SUBAPPLICATION AX_TO_QXA_BG_PUBLISH (* Treibt aus einem bereits fertigen AX-Zustand (z.B. per OR mehrerer Quellen zusammengefuehrt - gestaffeltes Gruppensignal, Einzel-Toggle, IO-Diag-Testbutton) 1 physischen Ausgang + Hintergrundfarbe (SoftKey+AUX) + lokalen State-Publish (Web-Client/OPC-Dashboard). Gegenstueck zu MyLib::sys::AX_SoftkeyToggle_RS_TO_QXA_BG (das den Toggle/Reset noch selbst erzeugt) - hier liegt der AX-Zustand bereits fertig vor und muss nur noch auf Ausgang+Hintergrund+Publish verteilt werden. *)
  (* Standard: 61499-2; Description: Copyright (c) 2026 Meisterschulen am Ostbahnhof This program and the accompanying materials are made available under the terms of the Eclipse Public License 2.0 which is available at https://www.eclipse.org/legal/epl-2.0/ SPDX-License-Identifier: EPL-2.0 *)
  (* Version 1.2, 2026-10-13, Franz Höpfinger, Meisterschulen am Ostbahnhof, Neuer SubAppEventOutput INITO (Type EInit), durchgereicht von DigitalOutput.INITO - analog ILOCK_SWITCH_2_QXA_OPC v1.3, fuer die Option-Lib-Migration Igel/Elevator Klassisch (echtes INIT_CNF statt T#15s-Delay-Raten). *)
  (* Version 1.1, 2026-10-12, Franz Höpfinger, Meisterschulen am Ostbahnhof, Neuer InputVar QI (BOOL) + SubAppEventInput INIT (Type EInit), durchgereicht an DigitalOutput.QI/.INIT statt hartem TRUE/Auto-Verteilung - QI-Gate Igel/Elevator Klassisch-vs-PVEA (gemeinsame Q5/Q7-Pins), 'Init wie bei Tecu'. Blast radius: 3 Instanzen, alle in Baender_EinAus.SUB (ueber AX_TO_QXA_BG_PUBLISH_SWITCHPIC) - bekommen alle ein explizites INIT statt Auto-Verteilung, unveraendertes Boot-Verhalten fuer Querband (sofort), neue Delay-Option fuer Igel/Elevator. *)
  PACKAGE MyLib::sys;
  IMPORT isobus::UT::Q::const::IDs::ID_NULL;
  IMPORT logiBUS::io::DQ::logiBUS_DO;
  IMPORT logiBUS::io::DQ::logiBUS_DO_S;
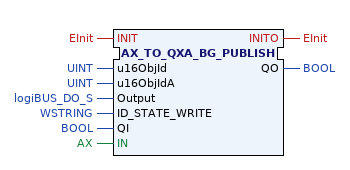
  EVENT_INPUT
    INIT : EInit; (* Initialisierung - durchgereicht an DigitalOutput.INIT statt Auto-Verteilung *)
  END_EVENT
  EVENT_OUTPUT
    INITO : EInit; (* Initialisierung abgeschlossen - echtes Confirm von DigitalOutput.INITO *)
  END_EVENT
  VAR_INPUT
    u16ObjId : UINT := ID_NULL; (* Object ID Softkey - traegt die Hintergrundfarbe *)
    u16ObjIdA : UINT := ID_NULL; (* Object ID AuxFunction2 (Joystick) - zeigt Hintergrundfarbe am Aux-Handle mit *)
    Output : logiBUS::io::DQ::logiBUS_DO_S := logiBUS_DO::Invalid; (* Identify the Output Output_Q1..Q12 *)
    ID_STATE_WRITE : WSTRING; (* Lokale Publish-Adresse (ACTION=WRITE) fuer den tatsaechlichen Zustand - wird von Web-Client/Dashboard remote abonniert *)
    QI : BOOL := TRUE; (* Qualifier fuer den physischen Ausgang - FALSE haelt diese Instanz komplett inaktiv *)
  END_VAR
  VAR_OUTPUT
    QO : BOOL; (* Quality Output - TRUE if service executed successfully (AND aus DigitalOutput/GreenWhiteBackground_AX/PUBLISH_STATE) *)
  END_VAR
  SOCKETS
    IN : adapter::types::unidirectional::AX; (* Fertiger AX-Zustand (bereits zusammengefuehrt) - wird auf Ausgang+Hintergrund+Publish verteilt *)
  END_SOCKETS
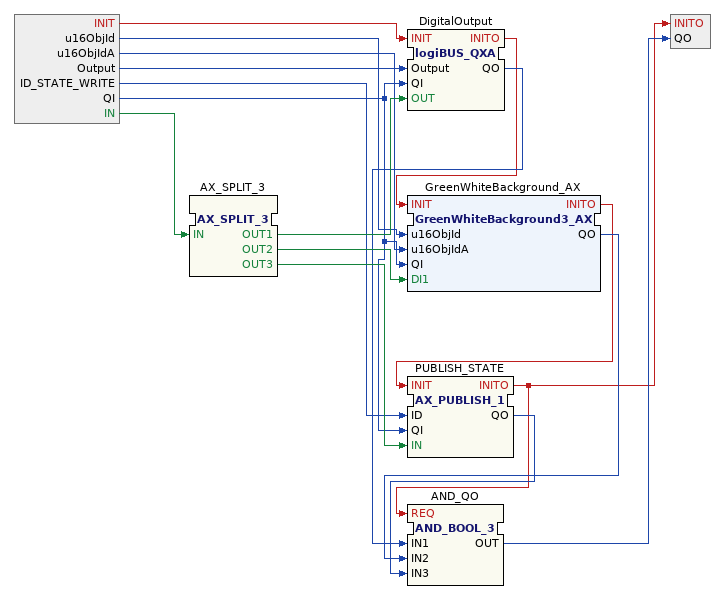
  FBS
    AX_SPLIT_3 : adapter::events::unidirectional::AX_SPLIT_3;
    DigitalOutput : logiBUS::io::DQ::logiBUS_QXA;
    PUBLISH_STATE : adapter::net::AX_PUBLISH_1;
    AND_QO : iec61131::booleanOperators::AND_BOOL_3;
  END_FBS
  SUBAPPS
    GreenWhiteBackground_AX : MyLib::sys::GreenWhiteBackground3_AX;
  END_SUBAPPS
  EVENT_CONNECTIONS
    INIT TO DigitalOutput.INIT;
    DigitalOutput.INITO TO GreenWhiteBackground_AX.INIT;
    GreenWhiteBackground_AX.INITO TO PUBLISH_STATE.INIT;
    PUBLISH_STATE.INITO TO INITO;
    PUBLISH_STATE.INITO TO AND_QO.REQ;
  END_CONNECTIONS
  DATA_CONNECTIONS
    u16ObjId TO GreenWhiteBackground_AX.u16ObjId;
    u16ObjIdA TO GreenWhiteBackground_AX.u16ObjIdA;
    Output TO DigitalOutput.Output;
    ID_STATE_WRITE TO PUBLISH_STATE.ID;
    QI TO DigitalOutput.QI;
    QI TO PUBLISH_STATE.QI;
    QI TO GreenWhiteBackground_AX.QI;
    DigitalOutput.QO TO AND_QO.IN1;
    GreenWhiteBackground_AX.QO TO AND_QO.IN2;
    PUBLISH_STATE.QO TO AND_QO.IN3;
    AND_QO.OUT TO QO;
  END_CONNECTIONS
  ADAPTER_CONNECTIONS
    IN TO AX_SPLIT_3.IN;
    AX_SPLIT_3.OUT1 TO DigitalOutput.OUT;
    AX_SPLIT_3.OUT2 TO GreenWhiteBackground_AX.DI1;
    AX_SPLIT_3.OUT3 TO PUBLISH_STATE.IN;
  END_CONNECTIONS
END_SUBAPPLICATION
